// CFC twin of T_SafeOpMode_Tests: the same tests drawn as CFC diagrams, the way a TwinSAFE project is authored.
    FUNCTION_BLOCK T_SafeOpMode_Tests_CFC EXTENDS T_SafeCfcTestSuite
    VAR
    // Test_ExactlyOneInputSelectsOutput
    group_1 : T_SafeGroup;
    fb_1 : T_SafeOpMode(group := group_1);
    // Test_ConnectedRestartRequiresRestartSequence
    group_2 : T_SafeGroup;
    fb_2 : T_SafeOpMode(group := group_2);
    // Test_SlowModeChangeGivesDiscrepancyError
    group_3 : T_SafeGroup;
    fb_3 : T_SafeOpMode(group := group_3) := (Parameters := (DiscrepancyTime := T#100MS));
    t0_3 : TON;
    t1_3 : TON;
    trig1_3 : R_TRIG;
END_VAR

Test_ExactlyOneInputSelectsOutput();
Test_ConnectedRestartRequiresRestartSequence();
Test_SlowModeChangeGivesDiscrepancyError();

METHOD PRIVATE Test_ExactlyOneInputSelectsOutput
// note: this text did not pass the execution check against the stored diagram
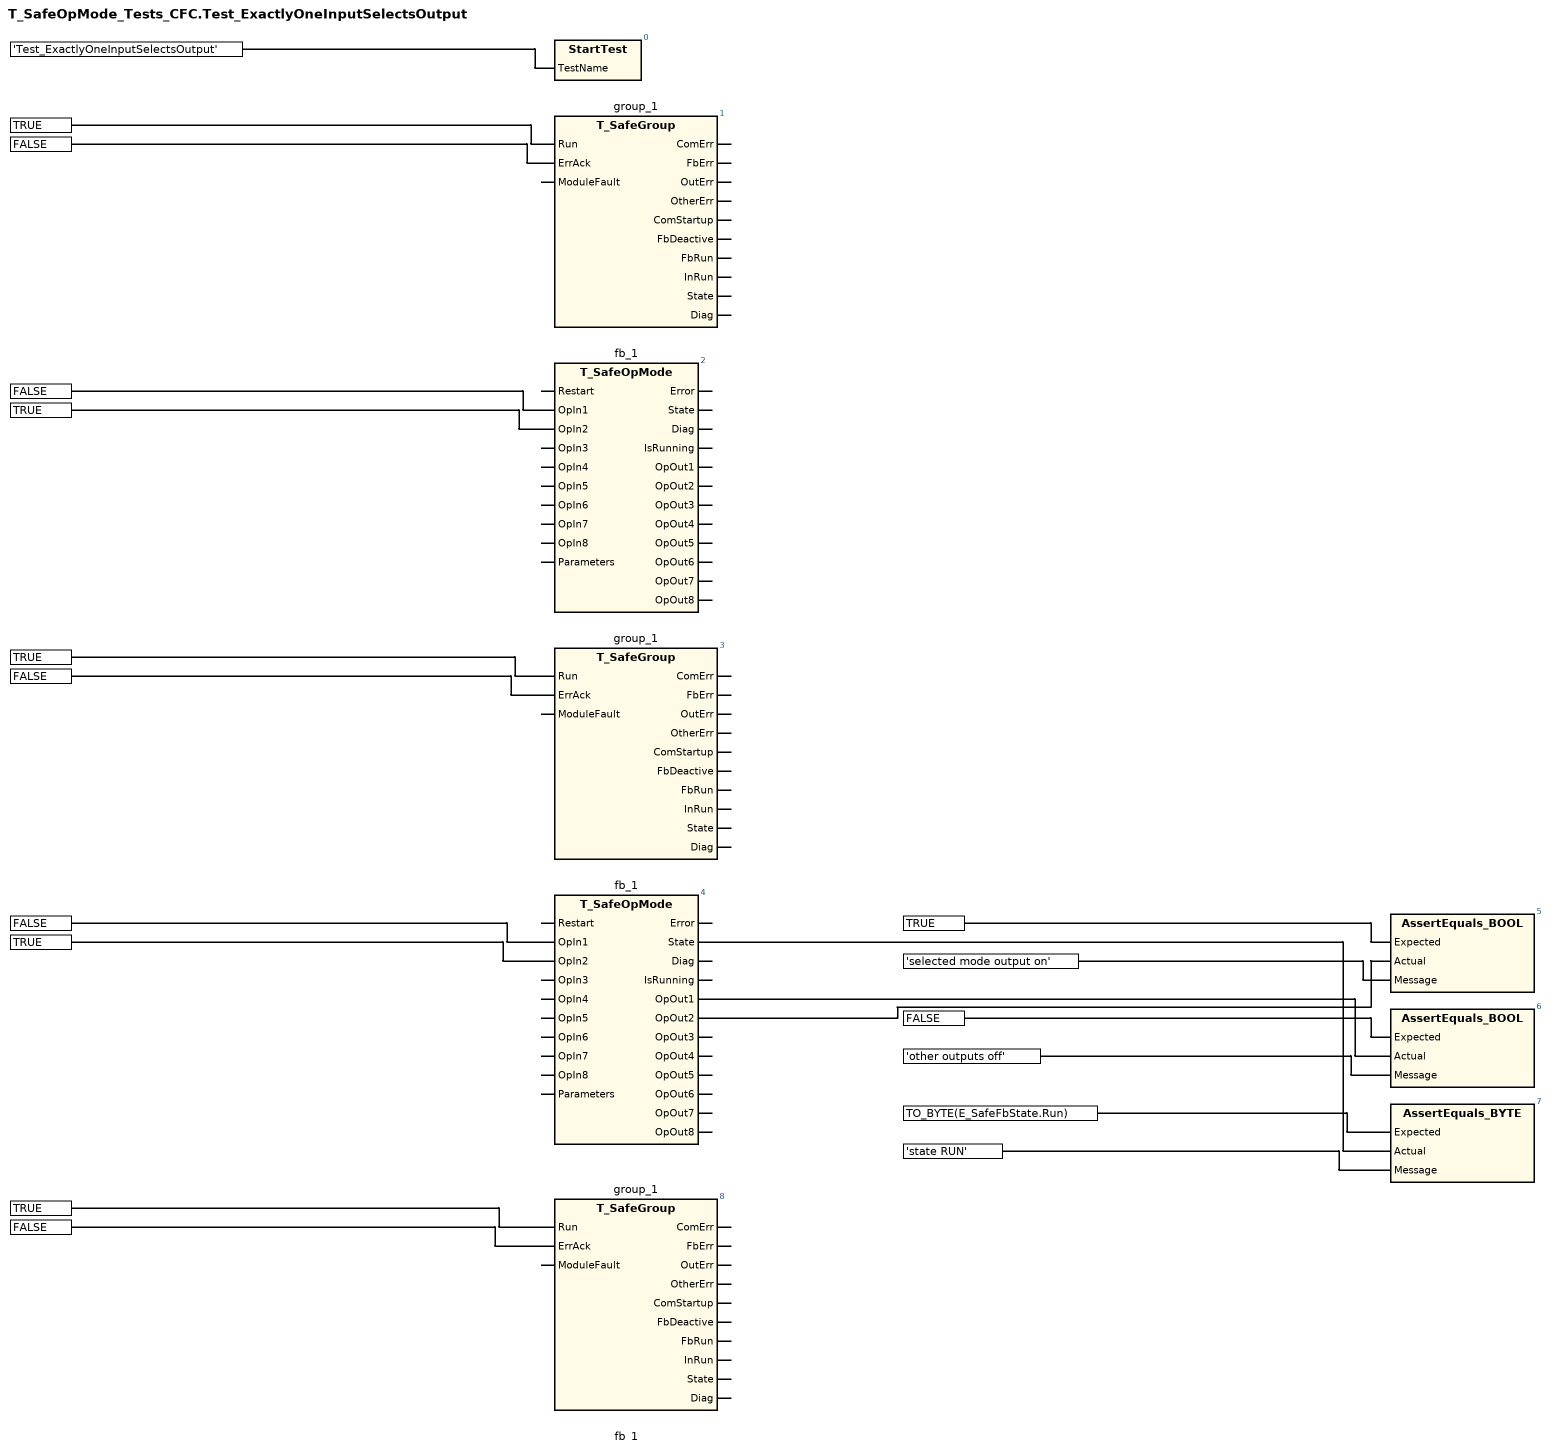
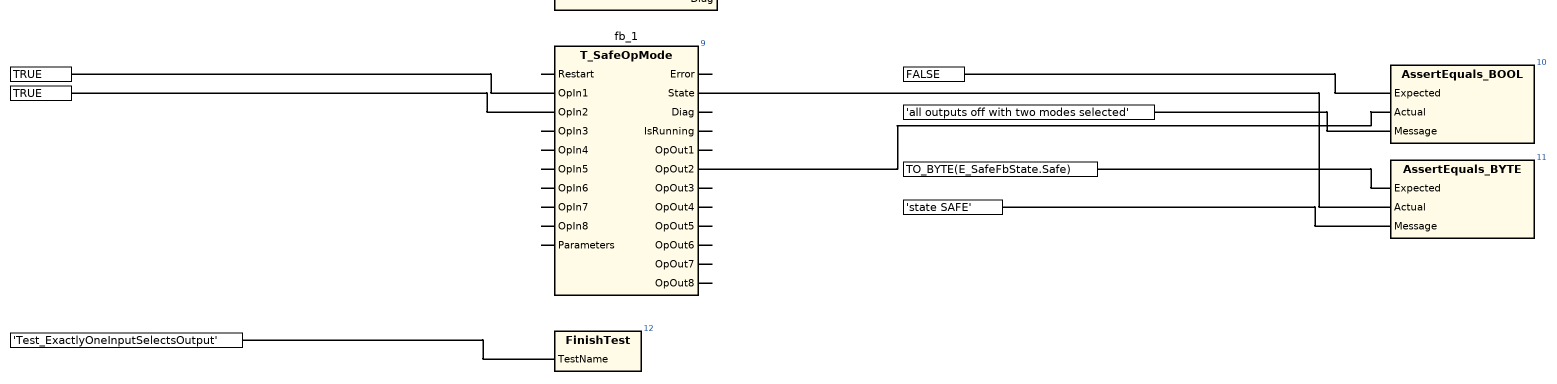
StartTest(TestName := 'Test_ExactlyOneInputSelectsOutput');
group_1(Run := TRUE, ErrAck := FALSE); // T_SafeGroup
fb_1(OpIn1 := FALSE, OpIn2 := TRUE); // T_SafeOpMode
group_1(Run := TRUE, ErrAck := FALSE); // T_SafeGroup
fb_1(OpIn1 := FALSE, OpIn2 := TRUE); // T_SafeOpMode
AssertEquals_BOOL(Expected := TRUE, Actual := fb_1.OpOut2, Message := 'selected mode output on');
AssertEquals_BOOL(Expected := FALSE, Actual := fb_1.OpOut1, Message := 'other outputs off');
AssertEquals_BYTE(Expected := TO_BYTE(E_SafeFbState.Run), Actual := fb_1.State, Message := 'state RUN');
group_1(Run := TRUE, ErrAck := FALSE); // T_SafeGroup
fb_1(OpIn1 := TRUE, OpIn2 := TRUE); // T_SafeOpMode
AssertEquals_BOOL(Expected := FALSE, Actual := fb_1.OpOut2, Message := 'all outputs off with two modes selected');
AssertEquals_BYTE(Expected := TO_BYTE(E_SafeFbState.Safe), Actual := fb_1.State, Message := 'state SAFE');
FinishTest(TestName := 'Test_ExactlyOneInputSelectsOutput');
END_METHOD

METHOD PRIVATE Test_ConnectedRestartRequiresRestartSequence
// note: this text did not pass the execution check against the stored diagram
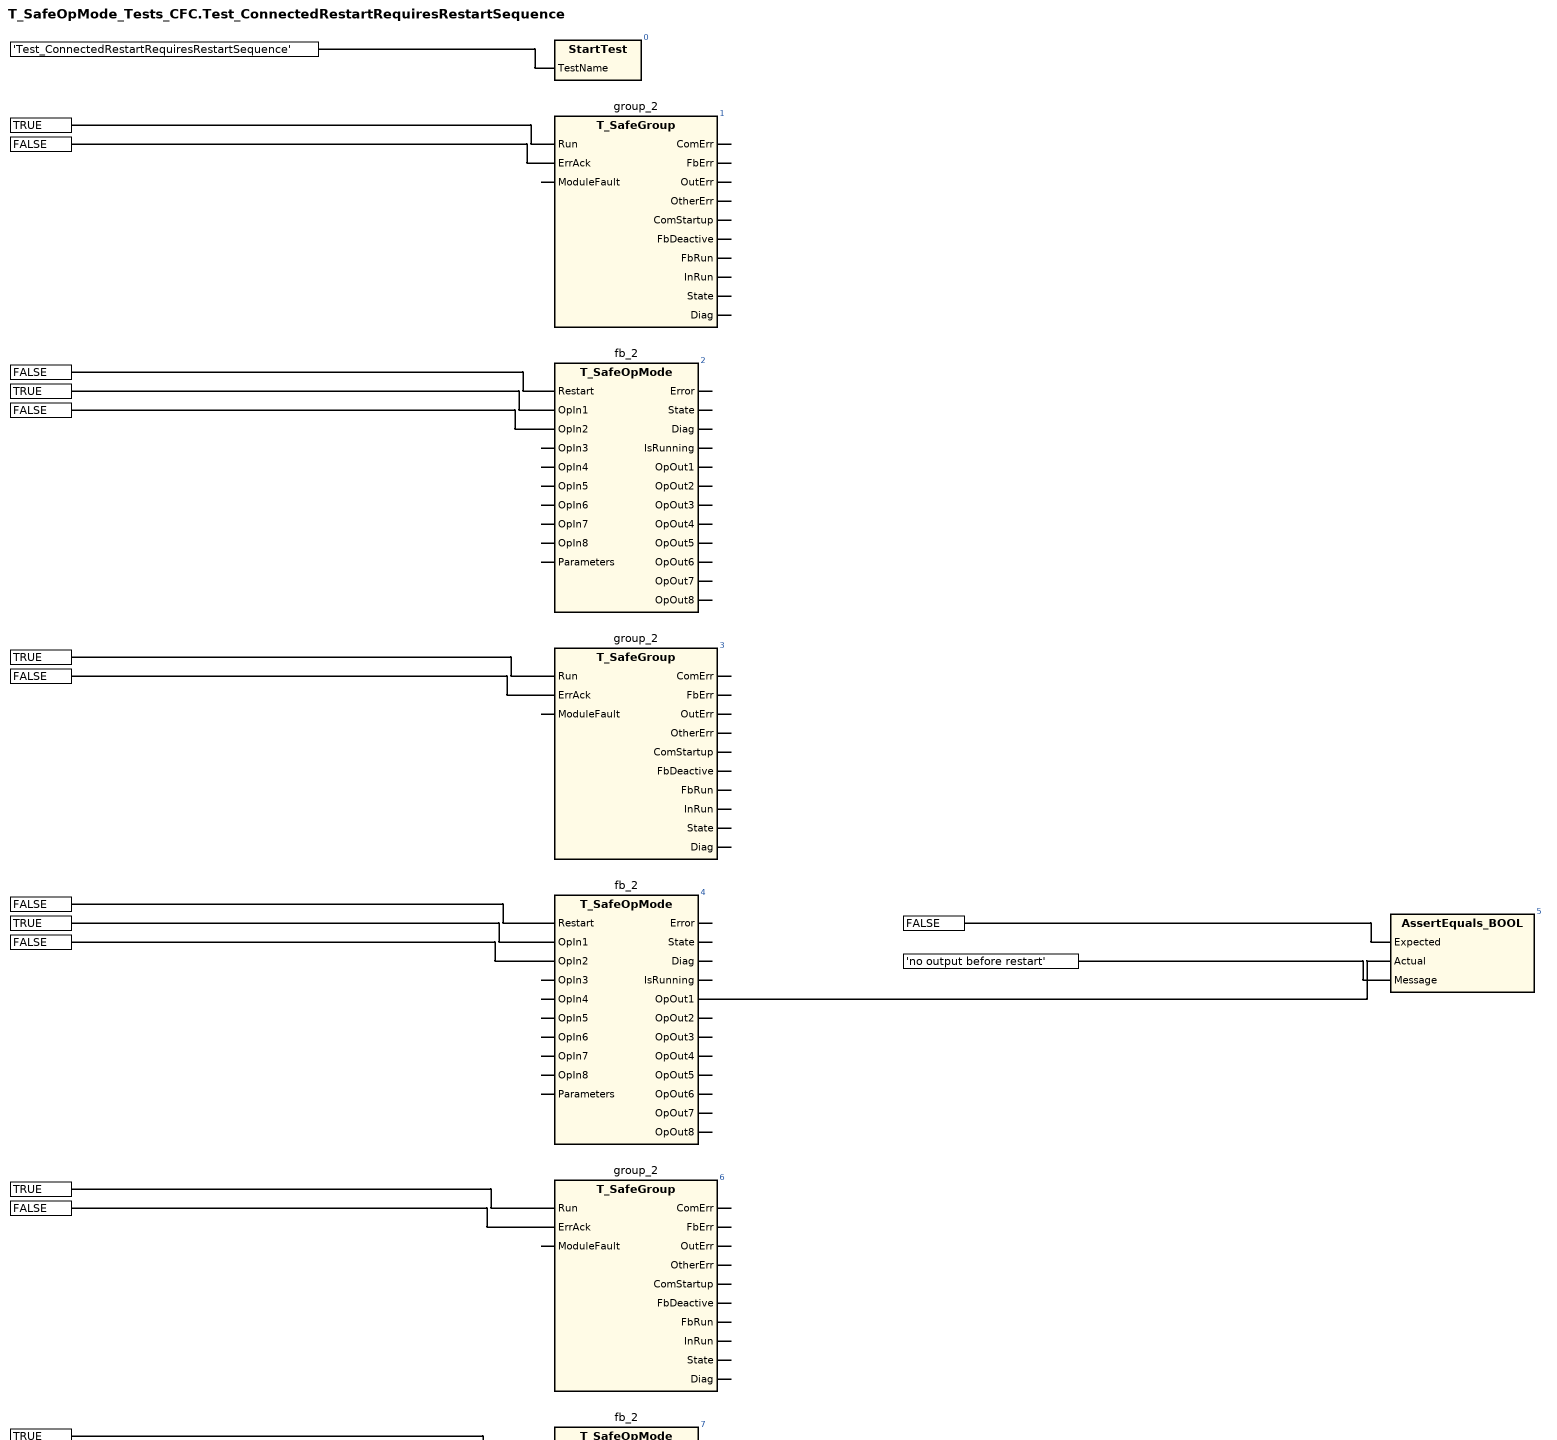
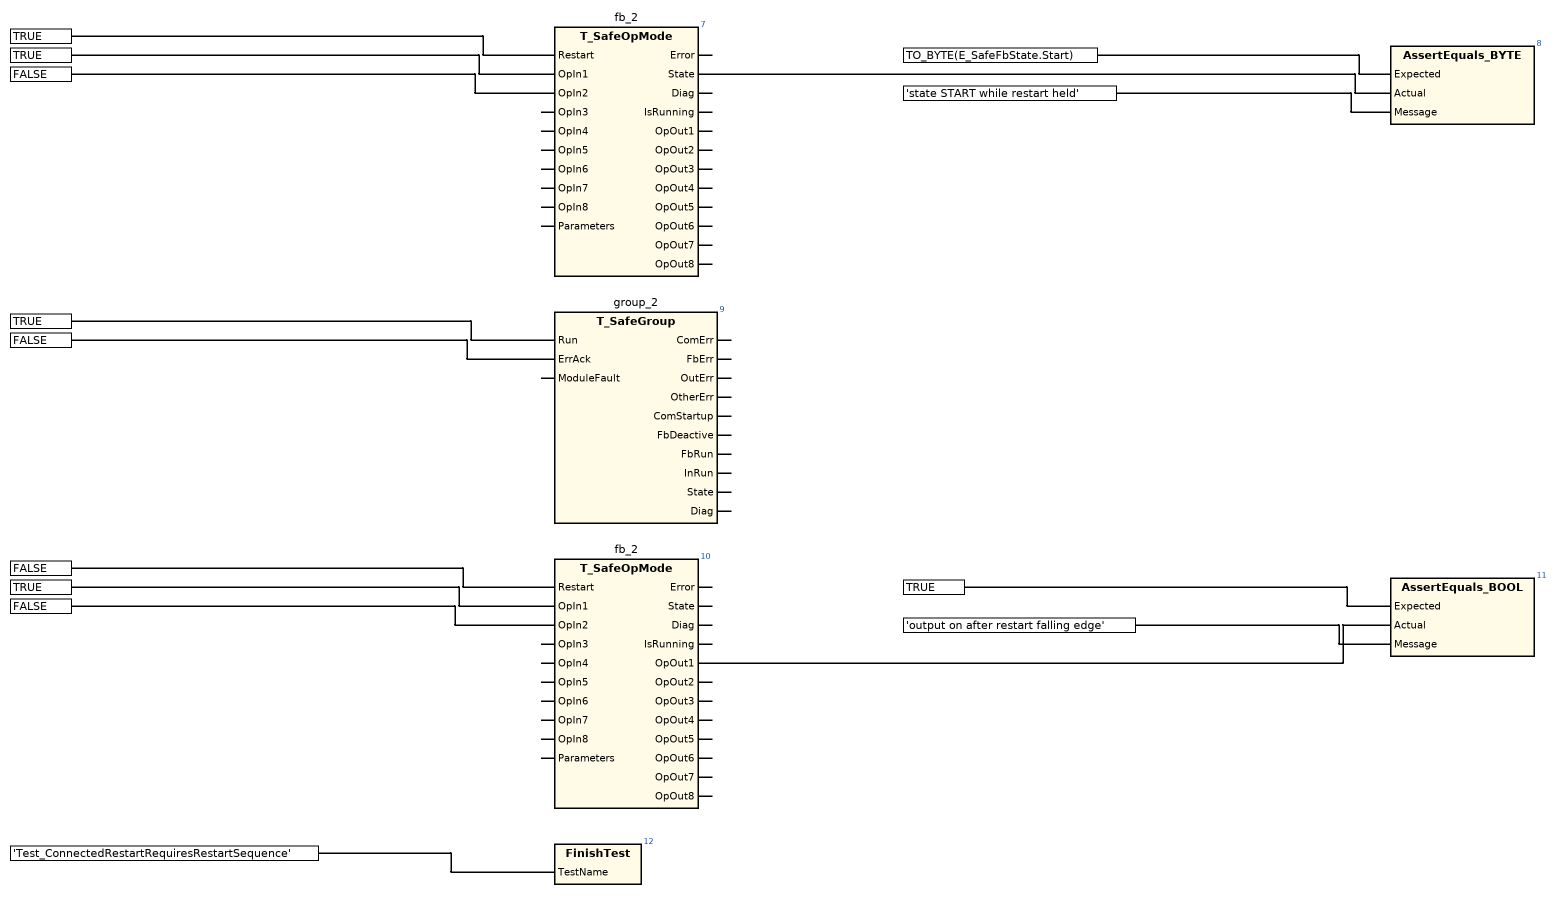
StartTest(TestName := 'Test_ConnectedRestartRequiresRestartSequence');
group_2(Run := TRUE, ErrAck := FALSE); // T_SafeGroup
fb_2(Restart := FALSE, OpIn1 := TRUE, OpIn2 := FALSE); // T_SafeOpMode
group_2(Run := TRUE, ErrAck := FALSE); // T_SafeGroup
fb_2(Restart := FALSE, OpIn1 := TRUE, OpIn2 := FALSE); // T_SafeOpMode
AssertEquals_BOOL(Expected := FALSE, Actual := fb_2.OpOut1, Message := 'no output before restart');
group_2(Run := TRUE, ErrAck := FALSE); // T_SafeGroup
fb_2(Restart := TRUE, OpIn1 := TRUE, OpIn2 := FALSE); // T_SafeOpMode
AssertEquals_BYTE(Expected := TO_BYTE(E_SafeFbState.Start), Actual := fb_2.State, Message := 'state START while restart held');
group_2(Run := TRUE, ErrAck := FALSE); // T_SafeGroup
fb_2(Restart := FALSE, OpIn1 := TRUE, OpIn2 := FALSE); // T_SafeOpMode
AssertEquals_BOOL(Expected := TRUE, Actual := fb_2.OpOut1, Message := 'output on after restart falling edge');
FinishTest(TestName := 'Test_ConnectedRestartRequiresRestartSequence');
END_METHOD

METHOD PRIVATE Test_SlowModeChangeGivesDiscrepancyError
// note: this text did not pass the execution check against the stored diagram
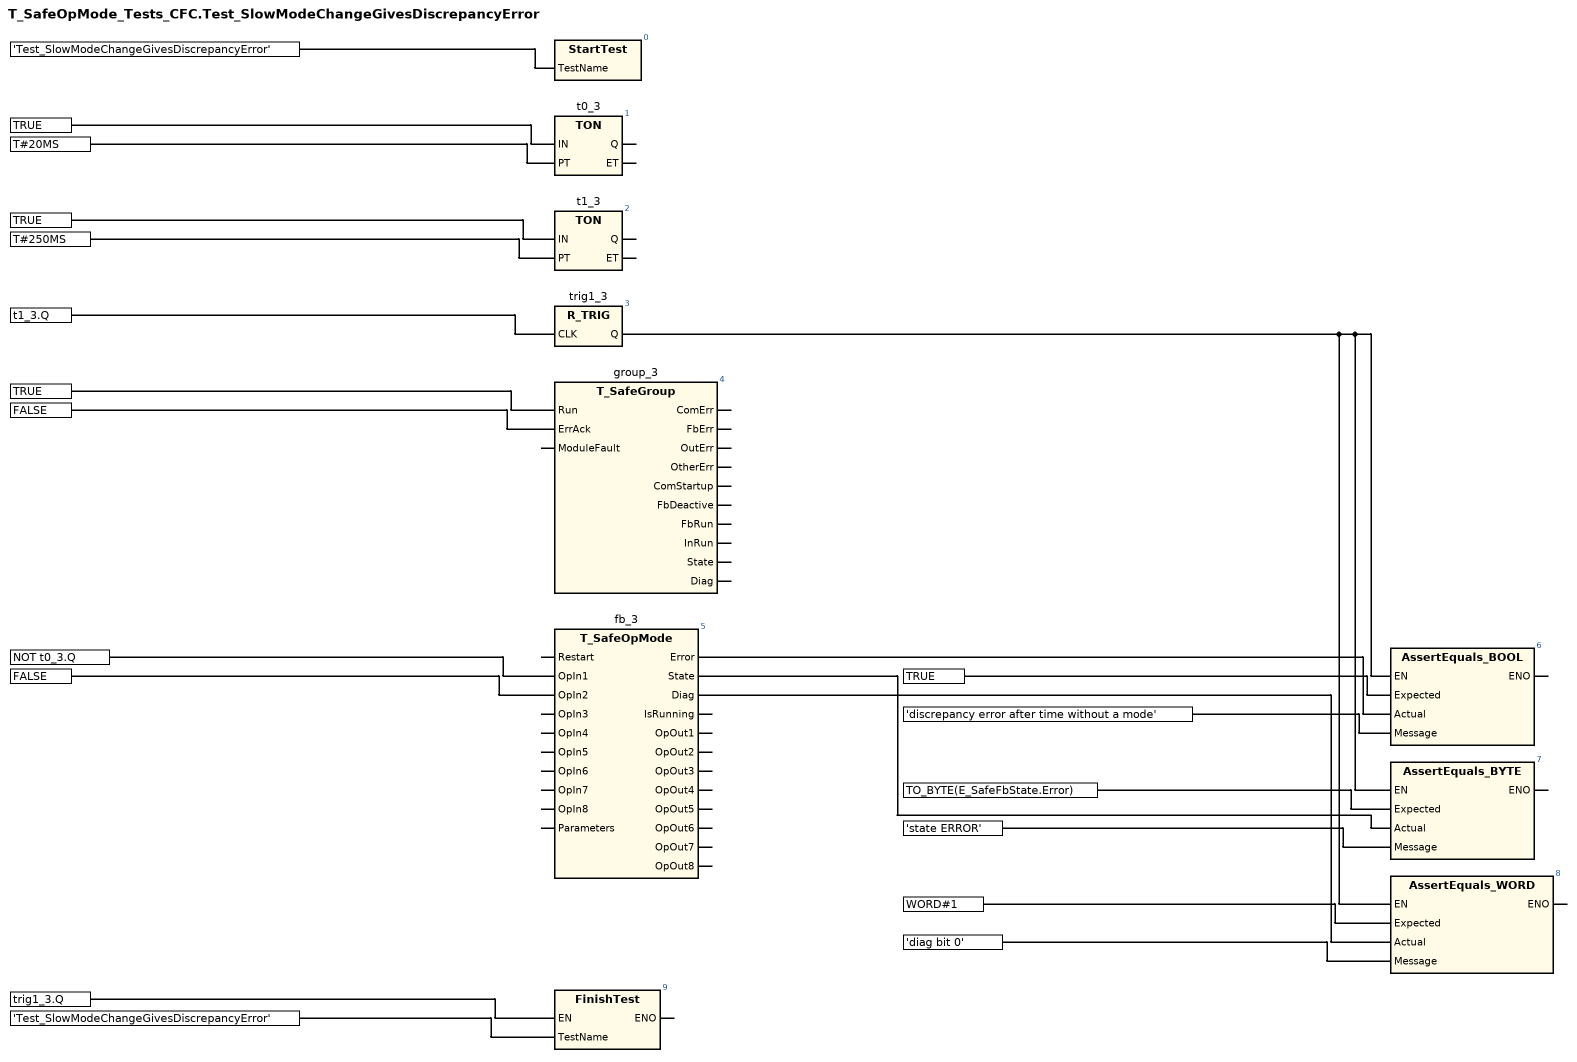
StartTest(TestName := 'Test_SlowModeChangeGivesDiscrepancyError');
t0_3(IN := TRUE, PT := T#20MS); // TON
t1_3(IN := TRUE, PT := T#250MS); // TON
trig1_3(CLK := t1_3.Q); // R_TRIG
group_3(Run := TRUE, ErrAck := FALSE); // T_SafeGroup
fb_3(OpIn1 := NOT t0_3.Q, OpIn2 := FALSE); // T_SafeOpMode
IF trig1_3.Q THEN AssertEquals_BOOL(Expected := TRUE, Actual := fb_3.Error, Message := 'discrepancy error after time without a mode'); END_IF
IF trig1_3.Q THEN AssertEquals_BYTE(Expected := TO_BYTE(E_SafeFbState.Error), Actual := fb_3.State, Message := 'state ERROR'); END_IF
IF trig1_3.Q THEN AssertEquals_WORD(Expected := WORD#1, Actual := fb_3.Diag, Message := 'diag bit 0'); END_IF
IF trig1_3.Q THEN FinishTest(TestName := 'Test_SlowModeChangeGivesDiscrepancyError'); END_IF
END_METHOD

END_FUNCTION_BLOCK

(* stored: Version 1.1.0.1, ProductVersion 3.1.4026.22
   POU T_SafeOpMode_Tests_CFC: Id {d4ff5807-e0e1-5d5f-bbc6-50a8a8e56b77}, SpecialFunc None
   Method Test_ExactlyOneInputSelectsOutput: Id {20910a78-aa36-5523-a359-fcbc1d508eb3}
   Method Test_ConnectedRestartRequiresRestartSequence: Id {370f51ab-d8d1-5a11-8da9-1940136e614d}
   Method Test_SlowModeChangeGivesDiscrepancyError: Id {30b83cfa-902d-5025-92ab-401d9a3afcb2} *)
